(* PLC project TBEN_L5_PLC11.project, CODESYS CODESYS V3.5 SP21 Patch 1 *)
(* stored: creationDateTime 2026-11-07T15:35:25.1897484, modificationDateTime 2026-11-07T15:09:07.4034196 *)

// Bố cục PDin O5D150 (16 bit, big-endian) - tách thành hằng để sửa theo IODD mà không đổi logic
TYPE ST_O5D150_PdLayout :
STRUCT
    usiOut1Bit       : USINT;      // bit OUT1 trong word PDin
    usiDistBitOffset : USINT;      // bit bắt đầu của Distance
    wDistMask        : WORD;       // mặt nạ sau khi dịch (12 bit = 16#0FFF)
    uiDistMin        : UINT;       // dải đo hợp lệ [cm]
    uiDistMax        : UINT;
    rGradient        : REAL;       // m / digit
END_STRUCT
END_TYPE
